(* CODESYS project BODAS-RC18-12_27-18_40-PAL.library
   Company: Bosch Rexroth AG
   DefaultNamespace: BODAS-API-RC18-12_27-18_40-PAL
   Title: BODAS_RC18-12_27-18_40-PAL
   DocFormat: reStructuredText
   Description: User library to use BODAS-BDL services (API) for RC40.
   Version: 2.3.0

Project tree, tasks and I/O mapping:
  PAL/
    API/
      function bds_snsrPal_getAgr [ST]
      function bds_snsrPal_getLnrPosn [ST]
    ENUM/
      data type bds_snsrPal_status_te
      data type bds_snsrPal_sigTyp_te
    STRUCT/
      data type bds_snsrPal_getLnrPosn_ts
      data type bds_snsrPal_getAgr_ts
      data type bds_snsrPalAnPwm_statusDiag_tb
      data type bds_snsrPalPwm_statusDiag_tb
      data type bds_snsrPalAn_statusDiag_tb
      data type bds_snsrPalSent_statusDiag_tb
    UNION/
      data type bds_snsrPal_statusDiag_tu
*)

// PAL/ENUM/bds_snsrPal_status_te
{attribute 'external_name' := 'cmp_rts_bds_snsrPal_status_te'}
TYPE bds_snsrPal_status_te :
(
    bds_snsrPal_ok_E := 0,                              // API call and function is ok
    bds_snsrPal_outOfRange_E := 1,                       // Detected Sensor Output1 and/or Sensor Output2 input values are out of range
    bds_snsrPal_outOfRangeErrOut2OkOut1_E := 2,         // Detected Sensor Output1 value is out of range and Sensor Output2 input value error
    bds_snsrPal_outOfRangeErrOut1OkOut2_E := 3,         // Detected Sensor Output1 input value error and Sensor Output1 input value is out of range
    bds_snsrPal_err_E := 4,                             // Sensor error detected or no data received
    bds_snsrPal_errMntd_E := 5,                         // Sensor magnet unit mounting error (magnet flux out of range 20-70mT)
    bds_snsrPal_errOut2OkOut1_E := 6,                   // Error on Sensor Output2 signal Sensor Output1 signal used for calculation
    bds_snsrPal_errOut1OkOut2_E := 7,                   // Error on Sensor Output1 signal Sensor Output2 signal used for calculation
    bds_snsrPal_invldConfig_E := 8,                     // Instance is not valid in active variant or not configured for the requested sensor
    bds_snsrPal_notConfig_E := 9,                       // Not configured e.g. RC4x Input1 and Input2 not configured for Sensor Output1 and Output2
    bds_snsrPal_invldPrm_E := 10                        // Wrong parameter
)USINT;
END_TYPE

// PAL/ENUM/bds_snsrPal_sigTyp_te
{attribute 'external_name' := 'cmp_rts_bds_snsrPal_sigTyp_te'}
TYPE bds_snsrPal_sigTyp_te :
(
    bds_snsrPalAnPwm_E := 0,                            // PAL analog and PWM sensor type
    bds_snsrPalAn_E := 1,                               // PAL analog sensor type
    bds_snsrPalPwm_E := 2,                              // PAL PWM sensor type
    bds_snsrPalSent_E := 3,                             // PAL SENT sensor type
    bds_snsrPalSigNotCfgd_E := 4                        // undefined sensor type
)USINT;
END_TYPE

// PAL/STRUCT/bds_snsrPal_getLnrPosn_ts
{attribute 'external_name' := 'cmp_bds_snsrPal_getLnrPosn_ts'}
TYPE bds_snsrPal_getLnrPosn_ts :
STRUCT
    stsApi_e: bds_snsrPal_status_te; //Return status information of API call
    sigTyp_e: bds_snsrPal_sigTyp_te; //Return status information of configured PAL sensor type for requested instance
    statusDiag_u: bds_snsrPal_statusDiag_tu; //Status diagnostic information of PAL sensor
    lnrPosn_uMtr_s32: DINT; //Measured linear position value from PAL sensor with resolution in micro meter
END_STRUCT
END_TYPE

// PAL/STRUCT/bds_snsrPal_getAgr_ts
{attribute 'external_name' := 'cmp_rts_bds_snsrPal_getAgr_ts'}
TYPE bds_snsrPal_getAgr_ts :
STRUCT
    stsApi_e: bds_snsrPal_status_te; //Return status information of API call
    sigTyp_e: bds_snsrPal_sigTyp_te; //Return status information of configured PAL sensor type for requested instance
    statusDiag_u: bds_snsrPal_statusDiag_tu; //Status diagnostic information of PAL sensor
    agr_mDeg_s32: DINT; //Measured angular value from PAL sensor with resolution in milli Degree
END_STRUCT
END_TYPE

// PAL/STRUCT/bds_snsrPalAnPwm_statusDiag_tb
{attribute 'external_name' := 'cmp_rts_bds_snsrPalAnPwm_statusDiag_tb'}
{attribute 'size' := '32'}
TYPE bds_snsrPalAnPwm_statusDiag_tb : STRUCT
    stLtdSfty1SigVal_b1 : BIT;          (* Fault error status bit information "Limited Safety" only one measured input signal value is valid or configured *)
    stLtdSftyCfgFlexInDev_b1 : BIT;     (* Fault error status bit information "Limited Safety" the two input signals are configured on the same FlexIn device *)
    stLtdSftyDeLim_b1 : BIT;            (* Fault error status bit information "Limited Safety" deviation of the measured input signal values above the limit value between the two input signals *)
    stErrAnSCB_b1 : BIT;                (* Fault error status for short cut to battery. TRUE: Short cut to battery is present. FALSE: Short cut to battery is not present *)
    stErrAnSCG_b1 : BIT;                (* Fault error status for short cut to ground. TRUE: Short cut to ground is present. FALSE: Short cut to ground is not present *)
    stErrAnOL_b1 : BIT;                 (* Fault error status for open load. TRUE: Open load is present. FALSE: Open load is not present *)
    stErrAnHw_b1 : BIT;                 (* Fault error status bit information of hardware error for analog voltage input. TRUE: Hardware error is present. FALSE: Hardware error is not present *)
    stErrPwmSnsr_b1 : BIT;              (* Fault error status bit information of sensor error for PWM input. TRUE: Sensor error is present. FALSE: Sensor error is not present *)
    stErrPwmHw_b1 : BIT;                (* Fault error status bit information of hardware error for PWM input. TRUE: Hardware error is present. FALSE: Hardware error is not present *)
    resd1_b : ARRAY[0..1] OF BYTE;      (* Reserved *)
END_STRUCT
END_TYPE

// PAL/UNION/bds_snsrPal_statusDiag_tu
{attribute 'external_name' := 'cmp_rts_bds_snsrPal_statusDiag_tu'}
TYPE bds_snsrPal_statusDiag_tu : UNION
    anPwmStDiag_b : bds_snsrPalAnPwm_statusDiag_tb;    (* Bit field for diagnostic information of PAL Analog/PWM sensor *)
    anStDiag_b : bds_snsrPalAn_statusDiag_tb;          (* Bit field for diagnostic information of PAL Analog/Analog sensor *)
    pwmStDiag_b : bds_snsrPalPwm_statusDiag_tb;        (* Bit field for diagnostic information of PAL PWM/PWM sensor *)
    sentStDiag_b : bds_snsrPalSent_statusDiag_tb;      (* Bit field for diagnostic information of PAL SENT/SENT sensor *)
    status_u32 : UDINT;                                (* General status bit diagnostic information of all PAL sensor interfaces *)
END_UNION
END_TYPE

// PAL/STRUCT/bds_snsrPalPwm_statusDiag_tb
{attribute 'external_name' := 'cmp_rts_bds_snsrPalPwm_statusDiag_tb'}
{attribute 'size' := '32'}
TYPE bds_snsrPalPwm_statusDiag_tb : STRUCT
    stLtdSfty1SigVal_b1 : BIT;          (* Fault error status bit information "Limited Safety" only one measured input signal value is valid or configured *)
    stLtdSftyCfgFlexInDev_b1 : BIT;     (* Fault error status bit information "Limited Safety" the two input signals are configured on the same FlexIn device *)
    stLtdSftyDeLim_b1 : BIT;            (* Fault error status bit information "Limited Safety" deviation of the measured input signal values above the limit value between the two input signals *)
    stErrPwm1Snsr_b1 : BIT;             (* Fault error status bit information for sensor error of PWM input 1. TRUE: Sensor error is present. FALSE: Sensor error is not present *)
    stErrPwm1Hw_b1 : BIT;               (* Fault error status bit information for hardware error of PWM input 1. TRUE: Hardware error is present. FALSE: Hardware error is not present *)
    stErrPwm2Snsr_b1 : BIT;             (* Fault error status bit information for sensor error of PWM input 2. TRUE: Sensor error is present. FALSE: Sensor error is not present *)
    stErrPwm2Hw_b1 : BIT;               (* Fault error status bit information for hardware error of PWM input 2. TRUE: Hardware error is present. FALSE: Hardware error is not present *)
    resd1_b : ARRAY[0..2] OF BYTE;      (* Unused bits *)
END_STRUCT
END_TYPE

// PAL/STRUCT/bds_snsrPalAn_statusDiag_tb
{attribute 'external_name' := 'cmp_rts_bds_snsrPalAn_statusDiag_tb'}
{attribute 'size' := '32'}
TYPE bds_snsrPalAn_statusDiag_tb : STRUCT
    stLtdSfty1SigVal_b1 : BIT;          (* Fault error status bit information "Limited Safety" only one measured input signal value is valid or configured *)
    stLtdSftyCfgFlexInDev_b1 : BIT;     (* Fault error status bit information "Limited Safety" the two input signals are configured on the same FlexIn device *)
    stLtdSftyDeLim_b1 : BIT;            (* Fault error status bit information "Limited Safety" deviation of the measured input signal values above the limit value between the two input signals *)
    stErrAn1SCB_b1 : BIT;               (* Fault error status bit information for short cut to battery of analog voltage input 1. TRUE: Short cut to battery is present. FALSE: Short cut to battery is not present *)
    stErrAn1SCG_b1 : BIT;               (* Fault error status bit information for short cut to ground of analog voltage input 1. TRUE: Short cut to ground is present. FALSE: Short cut to ground is not present *)
    stErrAn1OL_b1 : BIT;                (* Fault error status bit information for short cut to open load of analog voltage input 1. TRUE: Open load is present. FALSE: Open load is not present *)
    stErrAn1Hw_b1 : BIT;                (* Fault error status bit information for hardware error of analog voltage input 1. TRUE: Hardware error is present. FALSE: Hardware error is not present *)
    stErrAn2SCB_b1 : BIT;               (* Fault error status bit information for short cut to battery of analog voltage input 2. TRUE: Short cut to battery is present. FALSE: Short cut to battery is not present *)
    stErrAn2SCG_b1 : BIT;               (* Fault error status bit information for short cut to ground of analog voltage input 2. TRUE: Short cut to ground is present. FALSE: Short cut to ground is not present *)
    stErrAn2OL_b1 : BIT;                (* Fault error status bit information for short cut to open load of analog voltage input 2. TRUE: Open load is present. FALSE: Open load is not present *)
    stErrAn2Hw_b1 : BIT;                (* Fault error status bit information for hardware error of analog voltage input 2. TRUE: Hardware error is present. FALSE: Hardware error is not present *)
    resd1_b : ARRAY[0..1] OF BYTE;      (* Unused bits *)
END_STRUCT
END_TYPE

// PAL/STRUCT/bds_snsrPalSent_statusDiag_tb
{attribute 'external_name' := 'cmp_rts_bds_snsrPalSent_statusDiag_tb'}
{attribute 'size' := '32'}
TYPE bds_snsrPalSent_statusDiag_tb : STRUCT
    stLtdSfty1SigVal_b1 : BIT;              (* Fault error status bit information "Limited Safety" only one measured input signal value is valid or configured *)
    stLtdSftyCfgFlexInDev_b1 : BIT;         (* Fault error status bit information "Limited Safety" the two input signals are configured on the same FlexIn device *)
    stLtdSftyDeLim_b1 : BIT;                (* Fault error status bit information "Limited Safety" deviation for the measured input signal values above the limit value between the two input signals *)
    stErrSent1Snsr_b1 : BIT;                (* Fault error status bit information for angular or linear position above or below limit, overflows or saturation in supply voltage path (measurement possibly unreliable or wrong) or overflows or saturation in signal paths (pressure, temperature, supply voltage) for SENT input 1. TRUE: Sensor error is present. FALSE: Sensor error is not present *)
    stErrSent1Vdd_b1 : BIT;                 (* Fault error status bit information for low or high thresholds voltage supply exceeded of SENT input 1. TRUE: Sensor error is present. FALSE: Sensor error is not present *)
    stErrSent1Hw_b1 : BIT;                  (* Fault error status bit information for hardware error of SENT input 1. TRUE: Hardware error is present. FALSE: Hardware error is not present *)
    stErrSent1FldStrengthToHi_b1 : BIT;     (* Fault error status bit information for code field strength to high value error of SENT input 1. TRUE: Code field strength to high. FALSE: Code field strength in range *)
    stErrSent1FldStrengthToLo_b1 : BIT;     (* Fault error status bit information for code field strength to low value error of SENT input 1. TRUE: Code field strength to low. FALSE: Code field strength in range *)
    stErrSent1IvtMsn_b1 : BIT;              (* Fault error status bit information for inverted MSN data error of SENT input 1. TRUE: Inverted MSN data not match to SENT 1 position data. FALSE: Inverted MSN data match to SENT 1 position data *)
    stErrSent1SecaCntr_b1 : BIT;            (* Fault error status bit information for secure counter error of SENT input 1. TRUE: Secure counter is equal since last API function call. FALSE: Secure counter is unequal since last API function call *)
    stErrSent2Snsr_b1 : BIT;                (* Fault error status bit information for angular or linear position above or below limit, overflows or saturation in supply voltage path (measurement possibly unreliable or wrong) or overflows or saturation in signal paths (pressure, temperature, supply voltage) for SENT input 2. TRUE: Sensor error is present. FALSE: Sensor error is not present *)
    stErrSent2Vdd_b1 : BIT;                 (* Fault error status bit information for low or high thresholds voltage supply exceeded of SENT input 2. TRUE: Sensor error is present. FALSE: Sensor error is not present *)
    stErrSent2Hw_b1 : BIT;                  (* Fault error status bit information for hardware error of SENT input 2. TRUE: Hardware error is present. FALSE: Hardware error is not present *)
    stErrSent2FldStrengthToHi_b1 : BIT;     (* Fault error status bit information for code field strength to high value error of SENT input 2. TRUE: Code field strength to high. FALSE: Code field strength in range *)
    stErrSent2FldStrengthToLo_b1 : BIT;     (* Fault error status bit information for code field strength to low value error of SENT input 2. TRUE: Code field strength to low. FALSE: Code field strength in range *)
    resd1_b : ARRAY[0..1] OF BYTE;          (* Unused bits *)
END_STRUCT
END_TYPE

// PAL/API/bds_snsrPal_getAgr
/// The bds_snsrPal_getAgr API function provides the calculated angular position with resolution of milli-degree and diagnostic status of a PAL sensor instance.
///
///Remarks
///
/// The type of the sensor instance was configured in easyConfig.
/// If the function is called with an invalid PAL sensor instance or an error is detected, the function call status returns an error and the angular position value is set to 0x7FFFFFFF.
///
///Info
///
/// For safety-related application software, the “bit field” in the status diagnostic information of the PAL sensor “bds_snsrPal_statusDiag_tu statusDiag_u” must be checked by the customer to ensure that no safety bit
/// (stLtdSfty1SigVal_b1, stLtdSftyCfgFlexInDev_b1 and stLtdSftyDeLim_b1) is set to 1.
///
///==================================================================		  			===================================================================================================
///Return value    								  									     Description
///==================================================================		  			===================================================================================================
/// bds_snsrPal_getAgr_ts																 The return structure containing the status of the API function call, angular position in milli-degree and diagnostic information of the PAL sensor instance. For detail information please refer to chapter System feature BDL PAL 2/10.																	
///
///==================================================================		   			===================================================================================================
///
///=======
///Code Example:
///=======
///============================================================================
///
/// PROGRAM OsInitProc
///VAR
///
///    bds_snsrPal_getAgr_s : bds_snsrPal_getAgr_ts;
///	
///    bds_snsrPal_inst_e : bds_snsrPal_inst_te;
///	
///    agrLocal_mDeg_s32 : DINT := 75;
///	
///END_VAR
///
///bds_snsrPal_inst_e := bds_snsrPal_inst_te.PumpAngle_E;
///
///bds_snsrPal_getAgr_s := bds_snsrPal_getAgr(bds_snsrPal_inst_e);
///
/// (* check for safety application if return value can be used *)
/// IF bds_snsrPal_getAgr_s.stsApi_e = bds_snsrPal_ok_E THEN
///     (* check in return value if PAL PWM/Analog sensor type is configured *)
///     IF bds_snsrPal_getAgr_s.sigTyp_e = bds_snsrPalAnPwm_E THEN
///         (* error handling - check bit field status information of one signal is valid only *)
///         IF bds_snsrPal_getAgr_s.statusDiag_u.anPwmStDiag_b.stLtdSfty1SigVal_b1 = 1 THEN
///             (* usage of result only for none safety application software *)
///             (* ... *)
///             (* save the angular value in deci-degree from PAL sensor *)
///             agrLocal_mDeg_s32 := bds_snsrPal_getAgr_s.agr_mDeg_s32;
///         END_IF;
///         (* check bit field status information of detected Short Cut to Battery *)
///         IF bds_snsrPal_getAgr_s.statusDiag_u.anPwmStDiag_b.stErrAnSCB_b1 = 1 THEN
///             (* ... *)
///             (* save the angular value in deci-degree from PAL sensor *)
///             agrLocal_mDeg_s32 := 0;
///         END_IF;
///         (* ... *)
///     END_IF;
///     (* check in return value if PAL Analog/Analog sensor type is configured *)
///     IF bds_snsrPal_getAgr_s.sigTyp_e = bds_snsrPalAn_E THEN
///         (* ... *)
///     END_IF;
///     (* check also for PAL sensor types bds_snsrPalAn_E, bds_snsrPalPwm_E and bds_snsrPalSent_E *)
///     (* ... *)
/// ELSE
///     (* error handling *)
///     (* ... *)
/// END_IF;
/// END_PROGRAM
///
///============================================================================
{attribute 'external_name' := 'cmp_rts_bds_snsrPal_getAgr'}
FUNCTION bds_snsrPal_getAgr : bds_snsrPal_getAgr_ts
VAR_INPUT
    ///The PAL sensor instance name.
    snsrPalInst_e: USINT;
END_VAR

END_FUNCTION

// PAL/API/bds_snsrPal_getLnrPosn
/// The bds_snsrPal_getLnrPosn API function provides calculated linear position with resolution of micro-meter and diagnostic status of a PAL sensor instance.
///
///Remarks
///
/// The type of the sensor instance was configured in easyConfig.
/// If the function is called with an invalid PAL sensor instance or an error is detected, the function call status returns an error and the angular position value is set to 0x7FFFFFFF.
///
///  
///==================================================================		  			===================================================================================================
///Return value    								  									     Description
///==================================================================		  			===================================================================================================
/// bds_snsrPal_getLnrPosn_ts															The return structure containing the status of API function call, linear position in micro-meter and diagnostic information of a PAL sensor instance. For detail information please refer into chapter System feature BDL PAL 2/10.																
///
///==================================================================		   			===================================================================================================
///
///=======
///Code Example:
///=======
///============================================================================
///
/// PROGRAM OsInitProc
///VAR
///
///    bds_snsrPal_getLnrPosn_s : bds_snsrPal_getLnrPosn_ts;
///	
///    bds_snsrPal_inst_e : bds_snsrPal_inst_te;
///	
///    lnrPosnLocal_uMtr_s32 : DINT;
///	
///END_VAR
///
///bds_snsrPal_inst_e := bds_snsrPal_inst_te.PumpFrontRightLnrPosn_E;
///
///bds_snsrPal_getLnrPosn_s := bds_snsrPal_getLnrPosn(bds_snsrPal_inst_e);
///
/// IF(bds_snsrPal_ok_E = bds_snsrPal_getLnrPosn_s.stsApi_e) THEN
///         (* check in return value if PAL PWM/Analog sensor type is configured *)
///         IF bds_snsrPal_getLnrPosn_s.sigTyp_e = bds_snsrPalAnPwm_E THEN
///             (* error handling - check bit field status information of one signal is valid only *)
///             IF bds_snsrPal_getLnrPosn_s.statusDiag_u.anPwmStDiag_b.stLtdSfty1SigVal_b1 = 1 THEN
///                 (* usage of result only for none safety application software *)
///                 (* ... *)
///                 (* save the linear position value in micro-meter from PAL sensor *)
///                 lnrPosnLocal_uMtr_s32 := bds_snsrPal_getLnrPosn_s.lnrPosn_uMtr_s32;
///             END_IF;
///             (* check bit field status information of detected Short Cut to Battery *)
///             IF bds_snsrPal_getLnrPosn_s.statusDiag_u.anPwmStDiag_b.stErrAnSCB_b1 = 1 THEN
///                 (* ... *)
///                 (* save the angular value in milli-degree from PAL sensor *)
///                 lnrPosnLocal_uMtr_s32 := 0;
///             END_IF;
///             (* check all the other status information bits from bit field! *)
///             (* ... *)
///         END_IF;
///         (* check in return value if PAL Analog/Analog sensor type is configured *)
///         IF bds_snsrPal_getLnrPosn_s.sigTyp_e = bds_snsrPalAn_E THEN
///             (* ... *)
///         END_IF;
///         (* check also for PAL sensor types bds_snsrPalAn_E, bds_snsrPalPwm_E and bds_snsrPalSent_E *)
///         (* ... *)
/// ELSE
///     (* error handling *)
///     (* ... *)
/// END_IF;
/// END_PROGRAM
///
///============================================================================
{attribute 'external_name' := 'cmp_rts_bds_snsrPal_getLnrPosn'}
FUNCTION bds_snsrPal_getLnrPosn : bds_snsrPal_getLnrPosn_ts
VAR_INPUT
    ///The PAL sensor instance name.
    snsrPalInst_e: USINT;
END_VAR

END_FUNCTION
